// TwinCAT 3 PLC project PLCSim
// ProgramVersion: 3.1.4026.20
// libraries:
//   CmpBitmapPool, * (System)
//   Tc2_Standard, * (Beckhoff Automation GmbH)
//   Tc2_System, * (Beckhoff Automation GmbH)
//   Tc3_Module, * (Beckhoff Automation GmbH)
// project tree:
//   / GlobalTextList.TcGTLO, PlcTask.TcTTO, Visualization Manager.TcVMO (not stored)
//   GVLs/ GVL.TcGVL
//   POUs/ MAIN.TcPOU
//   VISUs/ ImagePool.TcIPO (not stored), Visualization.TcVIS
// real-time tasks:
//   TASK PlcTask: cycle T#80ms, priority 1, ADS port 350
//   TASK PlcTask1: cycle T#10ms, priority 20, ADS port 351
// variable links:
//   PLCSim/PLCSim Instance <-> PLCStudent/PLCStudent Instance
//     PlcTask Inputs/MAIN.ixRunConveyor1 <-> PlcTask Outputs/Control_FBD.qxRunConveyor1
//     PlcTask Inputs/MAIN.ixRunConveyor2 <-> PlcTask Outputs/Control_FBD.qxRunConveyor2
//     PlcTask Inputs/MAIN.ixRunConveyor3 <-> PlcTask Outputs/Control_FBD.qxRunConveyor3
//     PlcTask Outputs/MAIN.qxSensor1 <-> PlcTask Inputs/Control_FBD.ixSensor1
//     PlcTask Outputs/MAIN.qxSensor2 <-> PlcTask Inputs/Control_FBD.ixSensor2
//     PlcTask Outputs/MAIN.qxSensor3 <-> PlcTask Inputs/Control_FBD.ixSensor3

CONFIGURATION PLCSim
    RESOURCE PLC ON TwinCAT3
        TASK PlcTask(INTERVAL := T#80ms, PRIORITY := 1);
        PROGRAM MAIN WITH PlcTask : MAIN;
    END_RESOURCE
END_CONFIGURATION

// ---- GVLs/GVL.TcGVL
{attribute 'qualified_only'}
VAR_GLOBAL

END_VAR

// ---- POUs/MAIN.TcPOU
PROGRAM MAIN
VAR
	qxSensor1		AT %Q*:	BOOL; 		//Pallet on sensor1
	qxSensor2		AT %Q*:	BOOL; 		//Pallet on sensor2
	qxSensor3		AT %Q*:	BOOL; 		//Pallet on sensor3

	ixRunConveyor1	AT %I*:	BOOL; 		// Run Conveyor 1*)
	ixRunConveyor2	AT %I*:	BOOL; 		// Run Conveyor 2*)
	ixRunConveyor3	AT %I*:	BOOL; 		// Run Conveyor 3*)

	(* Internal Visiu variables *)
	miPallet1PosX:		INT:=0;		
	miPallet1PosY:		INT:=0;		
	miPallet2PosX:		INT:=0;	
	miPallet2PosY:		INT:=0;		
	miPallet3PosX:		INT:=0;
	miPallet3PosY:		INT:=0;		

	mxLoadPallet: BOOL;
	mxLoadPallet1: BOOL;
	mxLoadPallet2: BOOL;
	mxLoadPallet3: BOOL;
	
	mxMotor1Running : BOOL;
	mxMotor2Running : BOOL;
	mxMotor3Running : BOOL;
	
	mxEmptyConvayor1 : BOOL;
	mxEmptyConvayor2 : BOOL;
	mxEmptyConvayor3 : BOOL;
	
END_VAR

VAR CONSTANT

END_VAR

(*  Pallets on three conveyors  *)
(*  2024-10-29  Anders Nilsson University West *)


//Select a pallet to load
IF mxLoadPallet AND NOT qxSensor1 THEN
	IF miPallet1PosY = 0 AND NOT mxLoadPallet2 AND NOT mxLoadPallet3  THEN
		mxLoadPallet1 := TRUE;
	END_IF
	IF miPallet2PosY = 0 AND NOT mxLoadPallet1 AND NOT mxLoadPallet3  THEN
		mxLoadPallet2 := TRUE;
	END_IF
	IF miPallet3PosY = 0 AND NOT mxLoadPallet1 AND NOT mxLoadPallet2  THEN
		mxLoadPallet3 := TRUE;
	END_IF
END_IF
	
//Load Pallet 1	
IF mxLoadPallet1 THEN
	IF miPallet1PosY < 170 THEN 
		miPallet1PosY := miPallet1PosY + 5;
	ELSE 
		mxLoadPallet1 := FALSE;
	END_IF
END_IF

//Load Pallet 2	
IF mxLoadPallet2 THEN
	IF miPallet2PosY < 170 THEN 
		miPallet2PosY := miPallet2PosY + 5;
	ELSE 
		mxLoadPallet2 := FALSE;
	END_IF
END_IF

//Load Pallet 3	
IF mxLoadPallet3 THEN
	IF miPallet3PosY < 170 THEN 
		miPallet3PosY := miPallet3PosY + 5;
	ELSE 
		mxLoadPallet3 := FALSE;
	END_IF
END_IF

//Motor running signals to HMI
mxMotor1Running := ixRunConveyor1;
mxMotor2Running := ixRunConveyor2;
mxMotor3Running := ixRunConveyor3;


//Run Pallet 1 forward on conveyor 1
IF  ixRunConveyor1 AND miPallet1PosY = 170 AND miPallet1PosX < 120 THEN
	miPallet1PosX := miPallet1PosX + 2;
END_IF

//Run Pallet 1 forward on conveyor 2
IF  ixRunConveyor2 AND miPallet1PosY = 170 AND miPallet1PosX > 100 AND miPallet1PosX < 310 THEN
	miPallet1PosX := miPallet1PosX + 2;
END_IF

//Run Pallet 1 forward on conveyor 3
IF  ixRunConveyor3 AND miPallet1PosY = 170 AND miPallet1PosX > 290 AND miPallet1PosX < 500 THEN
	miPallet1PosX := miPallet1PosX + 2;
END_IF


//Run Pallet 2 forward on conveyor 1
IF  ixRunConveyor1 AND miPallet2PosY = 170 AND miPallet2PosX < 120 THEN
	miPallet2PosX := miPallet2PosX + 2;
END_IF

//Run Pallet 2 forward on conveyor 2
IF  ixRunConveyor2 AND miPallet2PosY = 170 AND miPallet2PosX > 100 AND miPallet2PosX < 310 THEN
	miPallet2PosX := miPallet2PosX + 2;
END_IF

//Run Pallet 2 forward on conveyor 3
IF  ixRunConveyor3 AND miPallet2PosY = 170 AND miPallet2PosX > 290 AND miPallet2PosX < 500 THEN
	miPallet2PosX := miPallet2PosX + 2;
END_IF

//Run Pallet 3 forward on conveyor 1
IF  ixRunConveyor1 AND miPallet3PosY = 170 AND miPallet3PosX < 120 THEN
	miPallet3PosX := miPallet3PosX + 2;
END_IF

//Run Pallet 3 forward on conveyor 2
IF  ixRunConveyor2 AND miPallet3PosY = 170 AND miPallet3PosX > 100 AND miPallet3PosX < 310 THEN
	miPallet3PosX := miPallet3PosX + 2;
END_IF

//Run Pallet 3 forward on conveyor 3
IF  ixRunConveyor3 AND miPallet3PosY = 170 AND miPallet3PosX > 290 AND miPallet3PosX < 500 THEN
	miPallet3PosX := miPallet3PosX + 2;
END_IF




//Empty the Pallets from conveyors
IF mxEmptyConvayor1 THEN 
	IF miPallet1PosY = 170 AND miPallet1PosX < 20 THEN
		miPallet1PosX := 0;
		miPallet1PosY := 0;
	END_IF
	IF miPallet2PosY = 170 AND miPallet2PosX < 20 THEN
		miPallet2PosX := 0;
		miPallet2PosY := 0;
	END_IF
	IF miPallet3PosY = 170 AND miPallet3PosX < 20 THEN
		miPallet3PosX := 0;
		miPallet3PosY := 0;
	END_IF
END_IF


IF mxEmptyConvayor2 THEN 
	IF miPallet1PosY = 170 AND miPallet1PosX >= 170 AND miPallet1PosX < 210   THEN
		miPallet1PosX := 0;
		miPallet1PosY := 0;
	END_IF
	IF miPallet2PosY = 170 AND miPallet2PosX >= 170 AND miPallet2PosX < 210 THEN
		miPallet2PosX := 0;
		miPallet2PosY := 0;
	END_IF
	IF miPallet3PosY = 170 AND miPallet3PosX >= 170 AND miPallet3PosX < 210 THEN
		miPallet3PosX := 0;
		miPallet3PosY := 0;
	END_IF	
	
END_IF

IF mxEmptyConvayor3 THEN
	IF miPallet1PosY = 170 AND miPallet1PosX >= 360 THEN 
		miPallet1PosX := 0;
		miPallet1PosY := 0;
	END_IF
	IF miPallet2PosY = 170 AND miPallet2PosX >= 360 THEN
		miPallet2PosX := 0;
		miPallet2PosY := 0;
	END_IF
	IF miPallet3PosY = 170 AND miPallet3PosX >= 360 THEN
		miPallet3PosX := 0;
		miPallet3PosY := 0;
	END_IF		
END_IF

//Sensors
qxSensor1 := miPallet1PosY = 170 AND miPallet1PosX < 150 
 		  OR miPallet2PosY = 170 AND miPallet2PosX < 150
		  OR miPallet3PosY = 170 AND miPallet3PosX < 150; 

qxSensor2 := miPallet1PosY = 170 AND miPallet1PosX > 200 AND miPallet1PosX < 330
          OR miPallet2PosY = 170 AND miPallet2PosX > 200 AND miPallet2PosX < 330
          OR miPallet3PosY = 170 AND miPallet3PosX > 200 AND miPallet3PosX < 330;

qxSensor3 := miPallet1PosY = 170 AND miPallet1PosX > 380 AND miPallet1PosX < 490
	      OR miPallet2PosY = 170 AND miPallet2PosX > 380 AND miPallet2PosX < 490
          OR miPallet3PosY = 170 AND miPallet3PosX > 380 AND miPallet3PosX < 490;

END_PROGRAM

// ---- GlobalTextList.TcGTLO
TEXTLIST GlobalTextList
  916 = '  LEVEL\nHIGHT                   NORM'
  815 = '  LEVEL\nNORM                   HIGH'
  391 = '  START                 STOP'
  77 = '  STOP                  START'
  297 = ' M1'
  505 = ' M2'
  534 = ' M3'
  5 = '%i'
  174 = '1'
  758 = '2'
  114 = '3'
  493 = 'ATM700 and ABD600 Exam 2025 '
  526 = 'CUR TEMP'
  6 = 'DISPLAY'
  143 = 'Empty Conveyor'
  951 = 'Empty Conveyor 1'
  288 = 'Empty Conveyor 2'
  559 = 'Empty Conveyor 3'
  176 = 'Exam 2025 ATM700 and ABD600 '
  417 = 'Exam 2025 in ATM700 and ABD600 '
  0 = 'Exam 2025, ATM700 and ABD600 '
  168 = 'Exam ATM700 and ABD600 '
  821 = 'LEVEL\nNORM                   HIGH'
  463 = 'Level 1'
  805 = 'Level 2'
  694 = 'Level 3'
  236 = 'Level Not Emty'
  86 = 'Load a pallet'
  87 = 'M1'
  227 = 'M2'
  462 = 'M3'
  142 = 'New pallet'
  825 = 'NORM '
  830 = 'Puls'
  172 = 'PULS'
  207 = 'Remove pallet'
  691 = 'S1'
  964 = 'S2'
  863 = 'S3'
  338 = 'Sensor 1'
  927 = 'Sensor 2'
  39 = 'Sensor 3'
  7 = 'SET TEMP'
  387 = 'STD200 Lab 1 '
  556 = 'Temp OK'
  910 = 'TEMP OK'
  215 = 'University West\nAnders N 2024'
  315 = 'University West\nAnders N 2025'
  141 = 'University West\nAnders N Dec 2018'
END_TEXTLIST

// ---- VISUs/Visualization.TcVIS
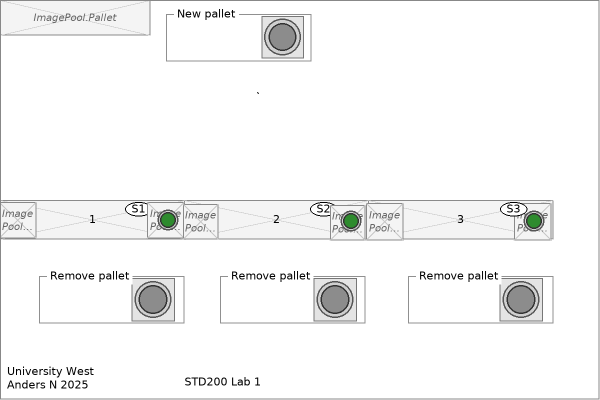
VISUALIZATION Visualization  // 600x400
    Label (4,363 125x30), "University West Anders N 2025"
    Image (0,200 185x39), "1", image: ImagePool.Conveyor
    Image (184,200 185x39), "2", image: ImagePool.Conveyor
    Image (368,200 185x39), "3", image: ImagePool.Conveyor
    Image (0,0 150x35), image: ImagePool.Pallet
        p3560616238: MAIN.miPallet1PosX
        p2738717112: MAIN.miPallet1PosY
    Image (0,0 150x35), image: ImagePool.Pallet
        p3560616238: MAIN.miPallet2PosX
        p2738717112: MAIN.miPallet2PosY
    Image (0,0 150x35), image: ImagePool.Pallet
        p3560616238: MAIN.miPallet3PosX
        p2738717112: MAIN.miPallet3PosY
    Image (514,203 37x37), invisible if: NOT MAIN.mxMotor3Running, image: ImagePool.Rotate
    Ellipse (125,202 27x14), "S1", tooltip "Sensor 1", colour toggle: MAIN.qxSensor1
    Ellipse (310,202 27x14), "S2", tooltip "Sensor 2", colour toggle: MAIN.qxSensor2
    Ellipse (500,202 27x14), "S3", tooltip "Sensor 3", colour toggle: MAIN.qxSensor3
    PushSwitch (497,278 48x43), tooltip "Empty Conveyor 3", variable: MAIN.mxEmptyConvayor3, behaviour: TAP, style: Switch-PushSwitch-Gray
    PushSwitch (311,278 48x43), tooltip "Empty Conveyor 2", variable: MAIN.mxEmptyConvayor2, behaviour: TAP, style: Switch-PushSwitch-Gray
    PushSwitch (129,278 48x43), tooltip "Empty Conveyor 1", variable: MAIN.mxEmptyConvayor1, behaviour: TAP, style: Switch-PushSwitch-Gray
    Image (-1,202 37x36), invisible if: NOT MAIN.mxMotor1Running, image: ImagePool.Rotate
    Image (147,202 37x36), invisible if: NOT MAIN.mxMotor1Running, image: ImagePool.Rotate
    Image (183,204 35x35), invisible if: NOT MAIN.mxMotor2Running, image: ImagePool.Rotate
    Image (330,205 35x35), invisible if: NOT MAIN.mxMotor2Running, image: ImagePool.Rotate
    Image (366,203 37x37), invisible if: NOT MAIN.mxMotor3Running, image: ImagePool.Rotate
    Label (99,363 251x38), "STD200 Lab 1"
    Polyline (257,92) (258,93)
    Lamp1 (155,208 26x24), variable: MAIN.mxMotor1Running, style: Lamp-Lamp1-Green
    Lamp1 (338,209 26x24), variable: MAIN.mxMotor2Running, style: Lamp-Lamp1-Green
    Lamp1 (521,209 26x24), variable: MAIN.mxMotor3Running, style: Lamp-Lamp1-Green
    Label (198,6 87x21)
    GroupBox (39,268 145x55), "Remove pallet"
    GroupBox (220,268 145x55), "Remove pallet"
    GroupBox (408,268 145x55), "Remove pallet"
    GroupBox (166,6 145x55), "New pallet"
        PushSwitch (94,10 45x42), tooltip "Load a pallet", variable: MAIN.mxLoadPallet, behaviour: TAP, style: Switch-PushSwitch-Gray
END_VISUALIZATION
